(* IEC 61131-3 sources: s7-to-codesys/tests/POUs/S7Compat/FB_S5Counter_Test, 5 files *)

(* ---- CountDownStopsAtZero.method.decl.st ---- *)
// CD уменьшает значение по фронту, но не ниже 0; A C = (значение <> 0).
METHOD PRIVATE CountDownStopsAtZero
VAR
    stCounter : ST_S5Counter;   // проверяемый счётчик
END_VAR

(* ---- CountUpOnEdgeUpTo999.method.decl.st ---- *)
// CU считает только фронты RLO; после установки 999 фронт CU значение не меняет.
METHOD PRIVATE CountUpOnEdgeUpTo999
VAR
    stCounter : ST_S5Counter;   // проверяемый счётчик (новый на каждый вызов метода)
END_VAR

(* ---- EnableRetriggersEdges.method.decl.st ---- *)
// FR C по фронту сбрасывает память фронтов: CU при удерживаемом RLO = 1 срабатывает снова; спад FR и
// удержание FR = 1 ничего не дают.
METHOD PRIVATE EnableRetriggersEdges
VAR
    stCounter : ST_S5Counter;   // проверяемый счётчик
END_VAR

(* ---- ResetIsLevel.method.decl.st ---- *)
// R C при RLO = 1 обнуляет значение на каждом вызове (по уровню), память фронтов не трогает.
METHOD PRIVATE ResetIsLevel
VAR
    stCounter : ST_S5Counter;   // проверяемый счётчик
END_VAR

(* ---- SetLoadsBcdOnEdge.method.decl.st ---- *)
// S C загружает BCD из ACCU1-L только по фронту; L C — двоичное значение, LC C — BCD.
METHOD PRIVATE SetLoadsBcdOnEdge
VAR
    stCounter : ST_S5Counter;   // проверяемый счётчик
END_VAR
